{region 'Documentation'}
(*!
<summary>Checks equality with the expected LTIME value.</summary>
*)
{endregion}
FUNCTION_BLOCK AssertEqual_LTime EXTENDS AssertionBase
VAR_INPUT
    IN : LTIME; //! Actual value checked or observed by this Assertion.
    Expected : LTIME; //! Reference value for comparison with IN.
END_VAR

SUPER^();

{region 'Documentation'}
(*!
<summary>Evaluate the typed duration relation and report higher-priority errors first.</summary>
*)
{endregion}
METHOD PROTECTED Assert
VAR
    Message : STRING(GVL_Constants.MessageLength);
    ExpectedText : STRING(GVL_Constants.AssertionValueLength);
    ActualText : STRING(GVL_Constants.AssertionValueLength);
END_VAR
IF NOT EvaluationActive THEN
    RETURN;
END_IF;

IF Result = E_Result.Error THEN
    RETURN;
END_IF;

IF Result = E_Result.Failed THEN
    RETURN;
END_IF;

IF IN <> Expected THEN
    ExpectedText := LTIME_TO_STRING(Expected);
    ActualText := LTIME_TO_STRING(IN);
    Message := CONCAT('Assertion failed: values are not equal. Expected = ',
        ExpectedText);
    Message := CONCAT(Message, ', Actual = ');
    Message := CONCAT(Message, ActualText);
    Message := CONCAT(Message, '.');
    Fail(Message := Message);
    RETURN;
END_IF;

Pass();
END_METHOD

END_FUNCTION_BLOCK

(* stored: Version 1.1.0.1
   POU AssertEqual_LTime: Id {76ae1a6f-07d4-463f-96ff-dbd7c5c660cd}, SpecialFunc None
   Folder Internal: Id {f171295f-ede5-4c0c-a145-5ceab86a8a8c}
   Method Assert: Id {c9af5bd4-038c-4123-9e17-2eab9fbd7cb4} *)
